# EPICS substitutions: apps/siemensApp/Db/bufdew_cpid.substitutions
file "db/siemens_cpid.db" {
pattern { P         PLCID       ORBV CVAL OVAL   MIN  MAX  DMIN  DMAX  VAL   KP   KI   KD  MDT  MMOD MVAL }
        { EV8210BP: PLC_BUFDEW  MD18 MD34 MD84  MD88 MD92 MD100 MD104 MD14  MD6 MD38 MD46 MD96 M42.0 MD50 }
        { EV8210:   PLC_BUFDEW  MD56 MD80 MD116 MD10 MD11 MD112 MD108 MD13 MD68 MD72 MD76 MD30 M64.0 MD60 }
}
